FUNCTION_BLOCK MOD_StateIds (* Builds the OPC UA addresses (Module/Reset ... Module/State) and the local channel names of the state manager. Technical: OPC UA and local channel IDs of the module state manager *)
  (* Standard: 61499-2 *)
  (* Version 0.1, 2026-09-28, Project contributors, AAU Smart Production Lab *)
  PACKAGE modlib;
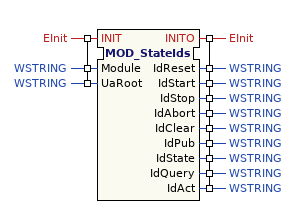
  EVENT_INPUT
    INIT : EInit WITH Module, UaRoot; (* Initialise, once at start-up (the INIT chain); takes the values given with it *)
  END_EVENT
  EVENT_OUTPUT
    INITO : EInit WITH IdReset, IdStart, IdStop, IdAbort, IdClear, IdPub, IdState, IdQuery, IdAct; (* Initialised: the next block of the INIT chain goes on *)
  END_EVENT
  VAR_INPUT
    Module : WSTRING; (* The module's name; its local channels are named after it (loc[<Module>/...]) *)
    UaRoot : WSTRING; (* The module's OPC UA folder, e.g. /Objects/Filling *)
  END_VAR
  VAR_OUTPUT
    IdReset : WSTRING; (* ID of the channel or OPC UA node of Reset *)
    IdStart : WSTRING; (* ID of the channel or OPC UA node of Start *)
    IdStop : WSTRING; (* ID of the channel or OPC UA node of Stop *)
    IdAbort : WSTRING; (* ID of the channel or OPC UA node of Abort *)
    IdClear : WSTRING; (* ID of the channel or OPC UA node of Clear *)
    IdPub : WSTRING; (* OPC UA ID of the published value *)
    IdState : WSTRING; (* Local channel of the module's state *)
    IdQuery : WSTRING; (* Local channel that asks for the current value (a block that starts later) *)
    IdAct : WSTRING; (* Local channel of the activity count *)
  END_VAR
  EC_STATES
    INIT : INIT -> INITO;
  END_STATES
  ALGORITHM INIT IN ST:
IdReset := CONCAT(CONCAT(CONCAT("opc_ua[CREATE_METHOD;", CONCAT(UaRoot, "/Module/")), "Reset"), "]");
IdStart := CONCAT(CONCAT(CONCAT("opc_ua[CREATE_METHOD;", CONCAT(UaRoot, "/Module/")), "Start"), "]");
IdStop := CONCAT(CONCAT(CONCAT("opc_ua[CREATE_METHOD;", CONCAT(UaRoot, "/Module/")), "Stop"), "]");
IdAbort := CONCAT(CONCAT(CONCAT("opc_ua[CREATE_METHOD;", CONCAT(UaRoot, "/Module/")), "Abort"), "]");
IdClear := CONCAT(CONCAT(CONCAT("opc_ua[CREATE_METHOD;", CONCAT(UaRoot, "/Module/")), "Clear"), "]");
IdPub := CONCAT(CONCAT(CONCAT("opc_ua[WRITE;", CONCAT(UaRoot, "/Module/")), "State"), "]");
IdState := CONCAT(CONCAT("loc[", Module), "/state]");
IdQuery := CONCAT(CONCAT("loc[", Module), "/state/query]");
IdAct := CONCAT(CONCAT("loc[", Module), "/activity]");
  END_ALGORITHM
END_FUNCTION_BLOCK
